Staubli VAL3: main.pgx

program main()
begin
  close(tCurrentTool)
  pPointRs.config.shoulder = lefty
  pPointRs2.config.shoulder = lefty
  mCurrentSpeed.tvel = 100.00
  mCurrentSpeed.blend = joint
  mCurrentSpeed.reach = 0.010
  mCurrentSpeed.leave = 0.010
  // Program TurnProg start
  // Program generated by RoboDK v6.0.7 for Staubli TP80 on XX/XX/XXXX 18:00:00
  // Using nominal kinematics.
  call MoveLine(-640.584,506.980,371.534,136.262,30.757,-130.375)
  call MoveLine(-607.850,543.849,363.215,136.262,30.757,-130.375)
  call MoveLine(-602.951,596.788,316.595,136.262,30.757,-130.375)
  pPointRs.config.shoulder = righty
  call MoveLine(-663.517,575.988,286.611,136.262,30.757,-130.375)
  pPointRs.config.shoulder = lefty
  call MoveLine(-650.861,503.437,361.399,136.262,30.757,-130.375)
  call MoveLine(-353.026,-90.135,331.702,164.619,39.324,-168.579)
  pPointRs.config.shoulder = righty
  call MoveLine(-624.230,571.208,454.620,81.604,51.756,-128.588)
  call MoveLine(-640.584,506.980,371.534,136.262,30.757,-130.375)
  call MoveJoint(350.00000,0.00000,0.00000,-350.00000)

  waitEndMove()
  // Program TurnProg end

end
